PROGRAM main
  VAR
    B1 AT %IX0.0  : BOOL; (* sensor de piezas *)
    S1 AT %IX0.1  : BOOL; (* RESET *)
    KM1 AT %QX0.0 : BOOL; (* motor de la cinta *)
    H1 AT %QX0.1  : BOOL; (* aviso *)
    PIEZAS        : CTU;
    CUENTA        : INT; (* piezas en la caja *)
  END_VAR

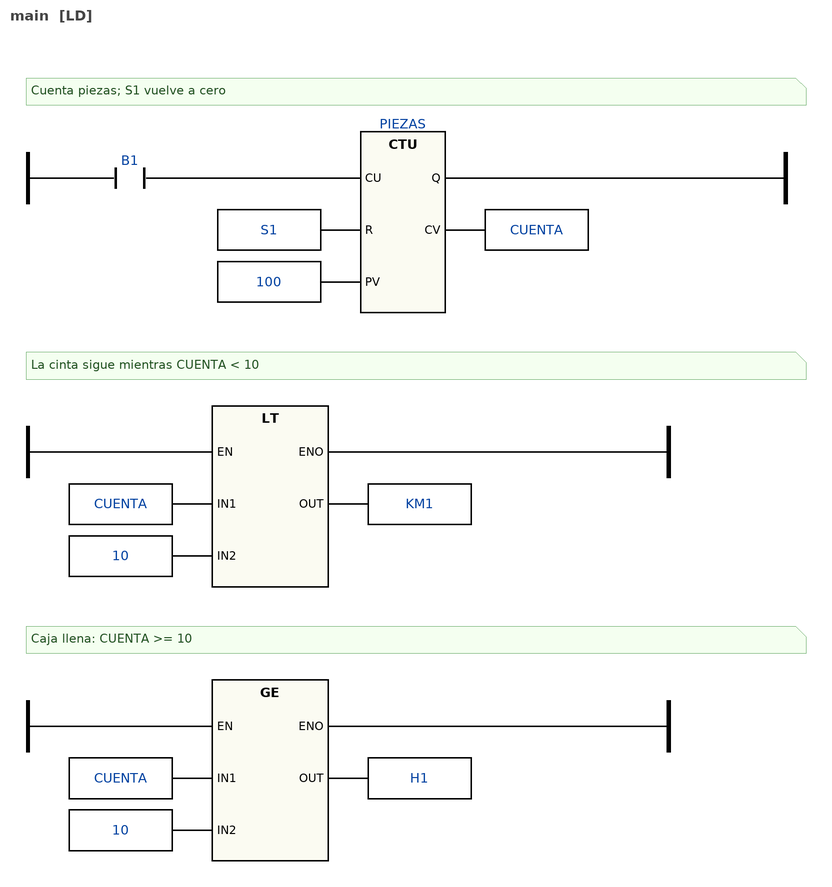
(* LD diagram, written out as Structured Text *)
(* Cuenta piezas; S1 vuelve a cero *)
PIEZAS(CU := B1, R := S1, PV := 100);
CUENTA := PIEZAS.CV;
(* La cinta sigue mientras CUENTA < 10 *)
KM1 := CUENTA < 10;
(* Caja llena: CUENTA >= 10 *)
H1 := CUENTA >= 10;
END_PROGRAM
